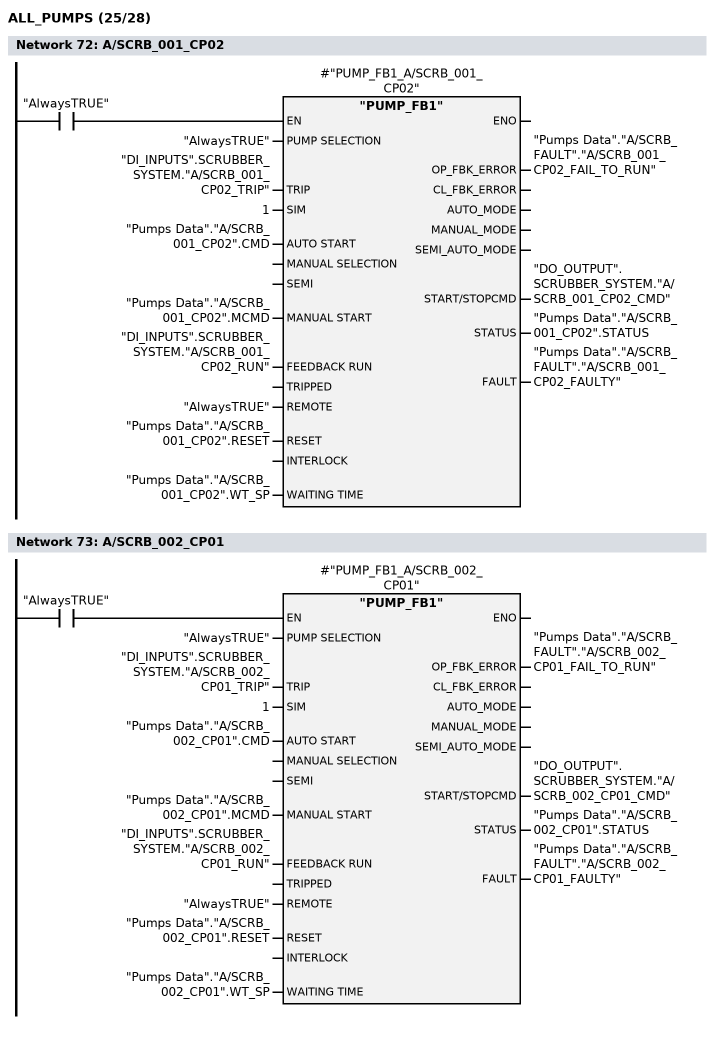
   RUNG wire#powerrail
      Contact( "AlwaysTRUE" )
      #"PUMP_FB1_A/SCRB_001_CP02"("PUMP SELECTION" := "AlwaysTRUE", TRIP := "DI_INPUTS".SCRUBBER_SYSTEM."A/SCRB_001_CP02_TRIP", SIM := 1, "AUTO START" := "Pumps Data"."A/SCRB_001_CP02".CMD, "MANUAL SELECTION" :=, SEMI :=, "MANUAL START" := "Pumps Data"."A/SCRB_001_CP02".MCMD, "FEEDBACK RUN" := "DI_INPUTS".SCRUBBER_SYSTEM."A/SCRB_001_CP02_RUN", TRIPPED :=, REMOTE := "AlwaysTRUE", RESET := "Pumps Data"."A/SCRB_001_CP02".RESET, INTERLOCK :=, "WAITING TIME" := "Pumps Data"."A/SCRB_001_CP02".WT_SP, OP_FBK_ERROR => "Pumps Data"."A/SCRB_FAULT"."A/SCRB_001_CP02_FAIL_TO_RUN", CL_FBK_ERROR =>, AUTO_MODE =>, MANUAL_MODE =>, SEMI_AUTO_MODE =>, "START/STOPCMD" => "DO_OUTPUT".SCRUBBER_SYSTEM."A/SCRB_001_CP02_CMD", STATUS => "Pumps Data"."A/SCRB_001_CP02".STATUS, FAULT => "Pumps Data"."A/SCRB_FAULT"."A/SCRB_001_CP02_FAULTY")
   END_RUNG
   // the same network as SCL:
   IF "AlwaysTRUE" THEN
       #"PUMP_FB1_A/SCRB_001_CP02"("PUMP SELECTION" := "AlwaysTRUE",   // "PUMP_FB1"
                               TRIP := "DI_INPUTS".SCRUBBER_SYSTEM."A/SCRB_001_CP02_TRIP",
                               SIM := 1,
                               "AUTO START" := "Pumps Data"."A/SCRB_001_CP02".CMD,
                               "MANUAL START" := "Pumps Data"."A/SCRB_001_CP02".MCMD,
                               "FEEDBACK RUN" := "DI_INPUTS".SCRUBBER_SYSTEM."A/SCRB_001_CP02_RUN",
                               REMOTE := "AlwaysTRUE",
                               RESET := "Pumps Data"."A/SCRB_001_CP02".RESET,
                               "WAITING TIME" := "Pumps Data"."A/SCRB_001_CP02".WT_SP,
                               OP_FBK_ERROR => "Pumps Data"."A/SCRB_FAULT"."A/SCRB_001_CP02_FAIL_TO_RUN",
                               "START/STOPCMD" => "DO_OUTPUT".SCRUBBER_SYSTEM."A/SCRB_001_CP02_CMD",
                               STATUS => "Pumps Data"."A/SCRB_001_CP02".STATUS,
                               FAULT => "Pumps Data"."A/SCRB_FAULT"."A/SCRB_001_CP02_FAULTY");
   END_IF;
END_REGION

REGION Network 73: A/SCRB_002_CP01
   RUNG wire#powerrail
      Contact( "AlwaysTRUE" )
      #"PUMP_FB1_A/SCRB_002_CP01"("PUMP SELECTION" := "AlwaysTRUE", TRIP := "DI_INPUTS".SCRUBBER_SYSTEM."A/SCRB_002_CP01_TRIP", SIM := 1, "AUTO START" := "Pumps Data"."A/SCRB_002_CP01".CMD, "MANUAL SELECTION" :=, SEMI :=, "MANUAL START" := "Pumps Data"."A/SCRB_002_CP01".MCMD, "FEEDBACK RUN" := "DI_INPUTS".SCRUBBER_SYSTEM."A/SCRB_002_CP01_RUN", TRIPPED :=, REMOTE := "AlwaysTRUE", RESET := "Pumps Data"."A/SCRB_002_CP01".RESET, INTERLOCK :=, "WAITING TIME" := "Pumps Data"."A/SCRB_002_CP01".WT_SP, OP_FBK_ERROR => "Pumps Data"."A/SCRB_FAULT"."A/SCRB_002_CP01_FAIL_TO_RUN", CL_FBK_ERROR =>, AUTO_MODE =>, MANUAL_MODE =>, SEMI_AUTO_MODE =>, "START/STOPCMD" => "DO_OUTPUT".SCRUBBER_SYSTEM."A/SCRB_002_CP01_CMD", STATUS => "Pumps Data"."A/SCRB_002_CP01".STATUS, FAULT => "Pumps Data"."A/SCRB_FAULT"."A/SCRB_002_CP01_FAULTY")
   END_RUNG
   // the same network as SCL:
   IF "AlwaysTRUE" THEN
       #"PUMP_FB1_A/SCRB_002_CP01"("PUMP SELECTION" := "AlwaysTRUE",   // "PUMP_FB1"
                               TRIP := "DI_INPUTS".SCRUBBER_SYSTEM."A/SCRB_002_CP01_TRIP",
                               SIM := 1,
                               "AUTO START" := "Pumps Data"."A/SCRB_002_CP01".CMD,
                               "MANUAL START" := "Pumps Data"."A/SCRB_002_CP01".MCMD,
                               "FEEDBACK RUN" := "DI_INPUTS".SCRUBBER_SYSTEM."A/SCRB_002_CP01_RUN",
                               REMOTE := "AlwaysTRUE",
                               RESET := "Pumps Data"."A/SCRB_002_CP01".RESET,
                               "WAITING TIME" := "Pumps Data"."A/SCRB_002_CP01".WT_SP,
                               OP_FBK_ERROR => "Pumps Data"."A/SCRB_FAULT"."A/SCRB_002_CP01_FAIL_TO_RUN",
                               "START/STOPCMD" => "DO_OUTPUT".SCRUBBER_SYSTEM."A/SCRB_002_CP01_CMD",
                               STATUS => "Pumps Data"."A/SCRB_002_CP01".STATUS,
                               FAULT => "Pumps Data"."A/SCRB_FAULT"."A/SCRB_002_CP01_FAULTY");
   END_IF;
END_REGION

REGION Network 74: A/SCRB_002_CP02
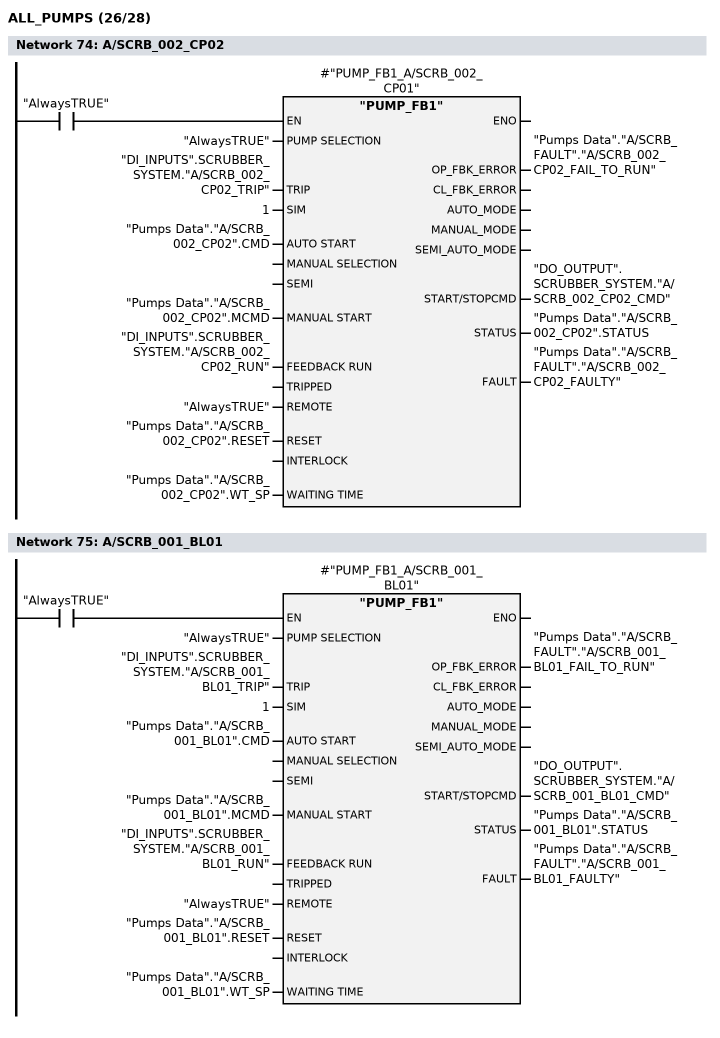
   RUNG wire#powerrail
      Contact( "AlwaysTRUE" )
      #"PUMP_FB1_A/SCRB_002_CP01"("PUMP SELECTION" := "AlwaysTRUE", TRIP := "DI_INPUTS".SCRUBBER_SYSTEM."A/SCRB_002_CP02_TRIP", SIM := 1, "AUTO START" := "Pumps Data"."A/SCRB_002_CP02".CMD, "MANUAL SELECTION" :=, SEMI :=, "MANUAL START" := "Pumps Data"."A/SCRB_002_CP02".MCMD, "FEEDBACK RUN" := "DI_INPUTS".SCRUBBER_SYSTEM."A/SCRB_002_CP02_RUN", TRIPPED :=, REMOTE := "AlwaysTRUE", RESET := "Pumps Data"."A/SCRB_002_CP02".RESET, INTERLOCK :=, "WAITING TIME" := "Pumps Data"."A/SCRB_002_CP02".WT_SP, OP_FBK_ERROR => "Pumps Data"."A/SCRB_FAULT"."A/SCRB_002_CP02_FAIL_TO_RUN", CL_FBK_ERROR =>, AUTO_MODE =>, MANUAL_MODE =>, SEMI_AUTO_MODE =>, "START/STOPCMD" => "DO_OUTPUT".SCRUBBER_SYSTEM."A/SCRB_002_CP02_CMD", STATUS => "Pumps Data"."A/SCRB_002_CP02".STATUS, FAULT => "Pumps Data"."A/SCRB_FAULT"."A/SCRB_002_CP02_FAULTY")
   END_RUNG
   // the same network as SCL:
   IF "AlwaysTRUE" THEN
       #"PUMP_FB1_A/SCRB_002_CP01"("PUMP SELECTION" := "AlwaysTRUE",   // "PUMP_FB1"
                               TRIP := "DI_INPUTS".SCRUBBER_SYSTEM."A/SCRB_002_CP02_TRIP",
                               SIM := 1,
                               "AUTO START" := "Pumps Data"."A/SCRB_002_CP02".CMD,
                               "MANUAL START" := "Pumps Data"."A/SCRB_002_CP02".MCMD,
                               "FEEDBACK RUN" := "DI_INPUTS".SCRUBBER_SYSTEM."A/SCRB_002_CP02_RUN",
                               REMOTE := "AlwaysTRUE",
                               RESET := "Pumps Data"."A/SCRB_002_CP02".RESET,
                               "WAITING TIME" := "Pumps Data"."A/SCRB_002_CP02".WT_SP,
                               OP_FBK_ERROR => "Pumps Data"."A/SCRB_FAULT"."A/SCRB_002_CP02_FAIL_TO_RUN",
                               "START/STOPCMD" => "DO_OUTPUT".SCRUBBER_SYSTEM."A/SCRB_002_CP02_CMD",
                               STATUS => "Pumps Data"."A/SCRB_002_CP02".STATUS,
                               FAULT => "Pumps Data"."A/SCRB_FAULT"."A/SCRB_002_CP02_FAULTY");
   END_IF;
END_REGION

REGION Network 75: A/SCRB_001_BL01
   RUNG wire#powerrail
      Contact( "AlwaysTRUE" )
      #"PUMP_FB1_A/SCRB_001_BL01"("PUMP SELECTION" := "AlwaysTRUE", TRIP := "DI_INPUTS".SCRUBBER_SYSTEM."A/SCRB_001_BL01_TRIP", SIM := 1, "AUTO START" := "Pumps Data"."A/SCRB_001_BL01".CMD, "MANUAL SELECTION" :=, SEMI :=, "MANUAL START" := "Pumps Data"."A/SCRB_001_BL01".MCMD, "FEEDBACK RUN" := "DI_INPUTS".SCRUBBER_SYSTEM."A/SCRB_001_BL01_RUN", TRIPPED :=, REMOTE := "AlwaysTRUE", RESET := "Pumps Data"."A/SCRB_001_BL01".RESET, INTERLOCK :=, "WAITING TIME" := "Pumps Data"."A/SCRB_001_BL01".WT_SP, OP_FBK_ERROR => "Pumps Data"."A/SCRB_FAULT"."A/SCRB_001_BL01_FAIL_TO_RUN", CL_FBK_ERROR =>, AUTO_MODE =>, MANUAL_MODE =>, SEMI_AUTO_MODE =>, "START/STOPCMD" => "DO_OUTPUT".SCRUBBER_SYSTEM."A/SCRB_001_BL01_CMD", STATUS => "Pumps Data"."A/SCRB_001_BL01".STATUS, FAULT => "Pumps Data"."A/SCRB_FAULT"."A/SCRB_001_BL01_FAULTY")
   END_RUNG
   // the same network as SCL:
   IF "AlwaysTRUE" THEN
       #"PUMP_FB1_A/SCRB_001_BL01"("PUMP SELECTION" := "AlwaysTRUE",   // "PUMP_FB1"
                               TRIP := "DI_INPUTS".SCRUBBER_SYSTEM."A/SCRB_001_BL01_TRIP",
                               SIM := 1,
                               "AUTO START" := "Pumps Data"."A/SCRB_001_BL01".CMD,
                               "MANUAL START" := "Pumps Data"."A/SCRB_001_BL01".MCMD,
                               "FEEDBACK RUN" := "DI_INPUTS".SCRUBBER_SYSTEM."A/SCRB_001_BL01_RUN",
                               REMOTE := "AlwaysTRUE",
                               RESET := "Pumps Data"."A/SCRB_001_BL01".RESET,
                               "WAITING TIME" := "Pumps Data"."A/SCRB_001_BL01".WT_SP,
                               OP_FBK_ERROR => "Pumps Data"."A/SCRB_FAULT"."A/SCRB_001_BL01_FAIL_TO_RUN",
                               "START/STOPCMD" => "DO_OUTPUT".SCRUBBER_SYSTEM."A/SCRB_001_BL01_CMD",
                               STATUS => "Pumps Data"."A/SCRB_001_BL01".STATUS,
                               FAULT => "Pumps Data"."A/SCRB_FAULT"."A/SCRB_001_BL01_FAULTY");
   END_IF;
END_REGION

REGION Network 76: A/SCRB_002_BL02
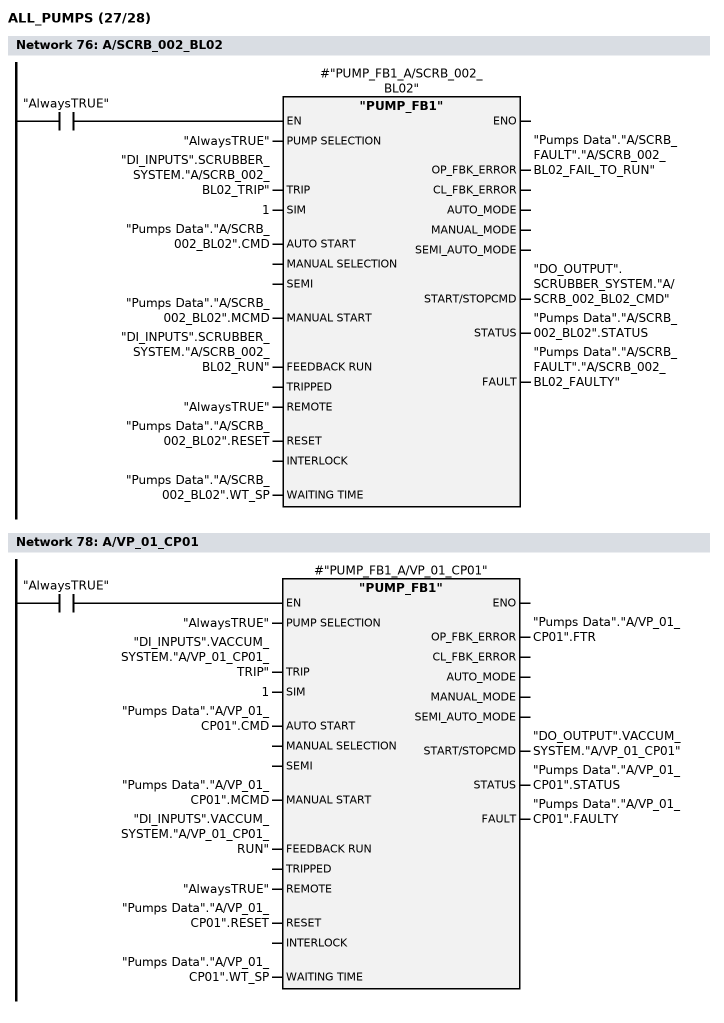
   RUNG wire#powerrail
      Contact( "AlwaysTRUE" )
      #"PUMP_FB1_A/SCRB_002_BL02"("PUMP SELECTION" := "AlwaysTRUE", TRIP := "DI_INPUTS".SCRUBBER_SYSTEM."A/SCRB_002_BL02_TRIP", SIM := 1, "AUTO START" := "Pumps Data"."A/SCRB_002_BL02".CMD, "MANUAL SELECTION" :=, SEMI :=, "MANUAL START" := "Pumps Data"."A/SCRB_002_BL02".MCMD, "FEEDBACK RUN" := "DI_INPUTS".SCRUBBER_SYSTEM."A/SCRB_002_BL02_RUN", TRIPPED :=, REMOTE := "AlwaysTRUE", RESET := "Pumps Data"."A/SCRB_002_BL02".RESET, INTERLOCK :=, "WAITING TIME" := "Pumps Data"."A/SCRB_002_BL02".WT_SP, OP_FBK_ERROR => "Pumps Data"."A/SCRB_FAULT"."A/SCRB_002_BL02_FAIL_TO_RUN", CL_FBK_ERROR =>, AUTO_MODE =>, MANUAL_MODE =>, SEMI_AUTO_MODE =>, "START/STOPCMD" => "DO_OUTPUT".SCRUBBER_SYSTEM."A/SCRB_002_BL02_CMD", STATUS => "Pumps Data"."A/SCRB_002_BL02".STATUS, FAULT => "Pumps Data"."A/SCRB_FAULT"."A/SCRB_002_BL02_FAULTY")
   END_RUNG
   // the same network as SCL:
   IF "AlwaysTRUE" THEN
       #"PUMP_FB1_A/SCRB_002_BL02"("PUMP SELECTION" := "AlwaysTRUE",   // "PUMP_FB1"
                               TRIP := "DI_INPUTS".SCRUBBER_SYSTEM."A/SCRB_002_BL02_TRIP",
                               SIM := 1,
                               "AUTO START" := "Pumps Data"."A/SCRB_002_BL02".CMD,
                               "MANUAL START" := "Pumps Data"."A/SCRB_002_BL02".MCMD,
                               "FEEDBACK RUN" := "DI_INPUTS".SCRUBBER_SYSTEM."A/SCRB_002_BL02_RUN",
                               REMOTE := "AlwaysTRUE",
                               RESET := "Pumps Data"."A/SCRB_002_BL02".RESET,
                               "WAITING TIME" := "Pumps Data"."A/SCRB_002_BL02".WT_SP,
                               OP_FBK_ERROR => "Pumps Data"."A/SCRB_FAULT"."A/SCRB_002_BL02_FAIL_TO_RUN",
                               "START/STOPCMD" => "DO_OUTPUT".SCRUBBER_SYSTEM."A/SCRB_002_BL02_CMD",
                               STATUS => "Pumps Data"."A/SCRB_002_BL02".STATUS,
                               FAULT => "Pumps Data"."A/SCRB_FAULT"."A/SCRB_002_BL02_FAULTY");
   END_IF;
END_REGION

REGION Network 78: A/VP_01_CP01
   RUNG wire#powerrail
      Contact( "AlwaysTRUE" )
      #"PUMP_FB1_A/VP_01_CP01"("PUMP SELECTION" := "AlwaysTRUE", TRIP := "DI_INPUTS".VACCUM_SYSTEM."A/VP_01_CP01_TRIP", SIM := 1, "AUTO START" := "Pumps Data"."A/VP_01_CP01".CMD, "MANUAL SELECTION" :=, SEMI :=, "MANUAL START" := "Pumps Data"."A/VP_01_CP01".MCMD, "FEEDBACK RUN" := "DI_INPUTS".VACCUM_SYSTEM."A/VP_01_CP01_RUN", TRIPPED :=, REMOTE := "AlwaysTRUE", RESET := "Pumps Data"."A/VP_01_CP01".RESET, INTERLOCK :=, "WAITING TIME" := "Pumps Data"."A/VP_01_CP01".WT_SP, OP_FBK_ERROR => "Pumps Data"."A/VP_01_CP01".FTR, CL_FBK_ERROR =>, AUTO_MODE =>, MANUAL_MODE =>, SEMI_AUTO_MODE =>, "START/STOPCMD" => "DO_OUTPUT".VACCUM_SYSTEM."A/VP_01_CP01", STATUS => "Pumps Data"."A/VP_01_CP01".STATUS, FAULT => "Pumps Data"."A/VP_01_CP01".FAULTY)
   END_RUNG
   // the same network as SCL:
   IF "AlwaysTRUE" THEN
       #"PUMP_FB1_A/VP_01_CP01"("PUMP SELECTION" := "AlwaysTRUE",   // "PUMP_FB1"
                               TRIP := "DI_INPUTS".VACCUM_SYSTEM."A/VP_01_CP01_TRIP",
                               SIM := 1,
                               "AUTO START" := "Pumps Data"."A/VP_01_CP01".CMD,
                               "MANUAL START" := "Pumps Data"."A/VP_01_CP01".MCMD,
                               "FEEDBACK RUN" := "DI_INPUTS".VACCUM_SYSTEM."A/VP_01_CP01_RUN",
                               REMOTE := "AlwaysTRUE",
                               RESET := "Pumps Data"."A/VP_01_CP01".RESET,
                               "WAITING TIME" := "Pumps Data"."A/VP_01_CP01".WT_SP,
                               OP_FBK_ERROR => "Pumps Data"."A/VP_01_CP01".FTR,
                               "START/STOPCMD" => "DO_OUTPUT".VACCUM_SYSTEM."A/VP_01_CP01",
                               STATUS => "Pumps Data"."A/VP_01_CP01".STATUS,
                               FAULT => "Pumps Data"."A/VP_01_CP01".FAULTY);
   END_IF;
END_REGION

REGION Network 79: A/VP_01_CP01
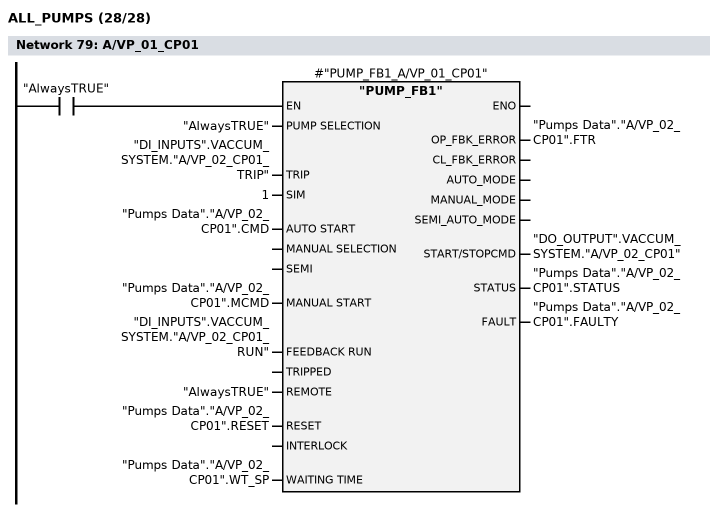
   RUNG wire#powerrail
      Contact( "AlwaysTRUE" )
      #"PUMP_FB1_A/VP_01_CP01"("PUMP SELECTION" := "AlwaysTRUE", TRIP := "DI_INPUTS".VACCUM_SYSTEM."A/VP_02_CP01_TRIP", SIM := 1, "AUTO START" := "Pumps Data"."A/VP_02_CP01".CMD, "MANUAL SELECTION" :=, SEMI :=, "MANUAL START" := "Pumps Data"."A/VP_02_CP01".MCMD, "FEEDBACK RUN" := "DI_INPUTS".VACCUM_SYSTEM."A/VP_02_CP01_RUN", TRIPPED :=, REMOTE := "AlwaysTRUE", RESET := "Pumps Data"."A/VP_02_CP01".RESET, INTERLOCK :=, "WAITING TIME" := "Pumps Data"."A/VP_02_CP01".WT_SP, OP_FBK_ERROR => "Pumps Data"."A/VP_02_CP01".FTR, CL_FBK_ERROR =>, AUTO_MODE =>, MANUAL_MODE =>, SEMI_AUTO_MODE =>, "START/STOPCMD" => "DO_OUTPUT".VACCUM_SYSTEM."A/VP_02_CP01", STATUS => "Pumps Data"."A/VP_02_CP01".STATUS, FAULT => "Pumps Data"."A/VP_02_CP01".FAULTY)
   END_RUNG
   // the same network as SCL:
   IF "AlwaysTRUE" THEN
       #"PUMP_FB1_A/VP_01_CP01"("PUMP SELECTION" := "AlwaysTRUE",   // "PUMP_FB1"
                               TRIP := "DI_INPUTS".VACCUM_SYSTEM."A/VP_02_CP01_TRIP",
                               SIM := 1,
                               "AUTO START" := "Pumps Data"."A/VP_02_CP01".CMD,
                               "MANUAL START" := "Pumps Data"."A/VP_02_CP01".MCMD,
                               "FEEDBACK RUN" := "DI_INPUTS".VACCUM_SYSTEM."A/VP_02_CP01_RUN",
                               REMOTE := "AlwaysTRUE",
                               RESET := "Pumps Data"."A/VP_02_CP01".RESET,
                               "WAITING TIME" := "Pumps Data"."A/VP_02_CP01".WT_SP,
                               OP_FBK_ERROR => "Pumps Data"."A/VP_02_CP01".FTR,
                               "START/STOPCMD" => "DO_OUTPUT".VACCUM_SYSTEM."A/VP_02_CP01",
                               STATUS => "Pumps Data"."A/VP_02_CP01".STATUS,
                               FAULT => "Pumps Data"."A/VP_02_CP01".FAULTY);
   END_IF;
END_REGION

REGION Network 80 (SCL)

   "A/SCRB_001_CP01_CMD" := "DO_OUTPUT".SCRUBBER_SYSTEM."A/SCRB_001_CP01_CMD";(*MODIFIED Q24.2 TO Q25.1*)
   "A/SCRB_001_CP02_CMD" := "DO_OUTPUT".SCRUBBER_SYSTEM."A/SCRB_001_CP02_CMD";
   "A/SCRB_001_BL01_CMD" := "DO_OUTPUT".SCRUBBER_SYSTEM."A/SCRB_001_BL01_CMD";
   "A/SCRB_002_CP01_CMD" := "DO_OUTPUT".SCRUBBER_SYSTEM."A/SCRB_002_CP01_CMD";
   "A/SCRB_002_CP02_CMD" := "DO_OUTPUT".SCRUBBER_SYSTEM."A/SCRB_002_CP02_CMD";
   "A/SCRB_002_BL01_CMD" := "DO_OUTPUT".SCRUBBER_SYSTEM."A/SCRB_002_BL02_CMD";
   "A/VP_01_CP01_CMD" := "DO_OUTPUT".VACCUM_SYSTEM."A/VP_01_CP01";
   "A/VP_02_CP01_CMD" := "DO_OUTPUT".VACCUM_SYSTEM."A/VP_02_CP01";
END_REGION
END_FUNCTION_BLOCK
